TYPE ST_PolarIIChamber_SingleProcessParam :
STRUCT
	ProcessStepCount : UINT; // 0..50; entries are contiguous from index 1
	ProcessSteps : ARRAY[1..50] OF ST_PolarIIChamber_ProcessStep;
	RecipeCount : UINT; // 0..50; entries are contiguous from index 1
	Recipes : ARRAY[1..50] OF ST_PolarIIChamber_Recipe;
END_STRUCT
END_TYPE

(* stored: Version 1.1.0.1, ProductVersion 3.1.4026.18
   DUT ST_PolarIIChamber_SingleProcessParam: Id {14000000-0000-0000-0000-000000000014} *)
